Staubli VAL3: main.pgx

program main()
begin
  close(tCurrentTool)
  pPointRx.config.shoulder = lefty
  pPointRx.config.elbow = epositive
  pPointRx.config.wrist = wpositive
  pPointRx2.config.shoulder = lefty
  pPointRx2.config.elbow = epositive
  pPointRx2.config.wrist = wpositive
  mCurrentSpeed.tvel = 100.00
  mCurrentSpeed.blend = joint
  mCurrentSpeed.reach = 0.010
  mCurrentSpeed.leave = 0.010
  // Program PrecProg start
  // Program generated by RoboDK v6.0.7 for Staubli RX130B on XX/XX/XXXX 18:00:00
  // Using nominal kinematics.
  call MoveJoint(12.34560,-45.67890,78.90130,-0.50000,0.49999,180.00000)
  call MoveLine(-640.585,506.981,371.534,136.641,31.137,-130.569)
  call MoveLine(0.500,-0.500,0.250,-180.000,0.005,-0.005)
  call MoveJoint(-12.34540,45.67850,-78.90000,0.50000,-0.00010,-180.00000)
  call MoveJoint(-12.34540,45.67850,-78.90000,0.50000,-0.00010,-180.00000)
  mCurrentSpeed.tvel = 66.667
  delay(0.002)
  delay(1.000)
  call MoveLine(-353.026,-90.135,331.702,164.619,39.324,-168.579)

  waitEndMove()
  // Program PrecProg end

end
